Fanuc KAREL source: ko00078.KL

-- PROVISIONAL review KL for V770-1; original PC SHA256 0fc7073be7c1220c855d122a8ea7357f4286afe85128f611f742601c90561083
-- Incomplete behavior may be omitted. Consult companion uncertainty JSON. Do not deploy.
PROGRAM KO00078
%NOLOCKGROUP
BEGIN
  -- UNRESOLVED_PC offsets 5-12; opcodes 9D,23
  -- UNRESOLVED_PC offsets 17-66; opcodes 27,22,1C,27,49,7E,AD,22,31,7E,4A
  -- UNRESOLVED_PC offsets 71-75; opcodes 7F
END KO00078
